(* IEC 61131-3 sources: krc-sample-programs/robot-cell-ethernetip-codesys/source/06_Programs, 5 files *)

(* ---- DASHBOARD.st ---- *)
PROGRAM DASHBOARD
VAR
	ipRobot      : NBS.IPv4Address := (ipAddress := ROBOT_IP);	// The robot's address
	fbClient     : NBS.TCP_Client;	// The connection to the robot's Dashboard Server
	fbWrite      : NBS.TCP_Write;	// Sends one line
	fbRead       : NBS.TCP_Read;	// Takes in whatever the robot has sent
	TON_POLL     : TON;	// Paces the questions
	TON_REPLY    : TON;	// The robot's answer is overdue
	TON_RETRY    : TON;	// Still not connected: try again
	bDropped     : BOOL;	// The connection was dropped this scan, so the retry timer starts over
	iDashStep    : INT;	// 0 not connected, 10 waiting for hello, 20 idle, 30 sending, 40 waiting for the answer
	bReconnect   : BOOL;	// Drop the connection for one scan, to connect again
	bAskRemote   : BOOL;	// The question in flight, or the next one, is remote control (the two take turns)
	sOut         : STRING(80);	// The line going out, with its line feed
	abIn         : ARRAY[0..127] OF BYTE;	// The bytes the read brings in
	sLine        : STRING(80);	// The line coming in, put together up to its line feed
	bLineDone    : BOOL;	// A whole line has come in this scan
	sChar        : STRING(1);	// One character, to add to the line
	i            : UDINT;	// Counts through the bytes read
END_VAR
// ---- body ----
// DASHBOARD: the driver for the second connection to the robot, its Dashboard Server. Not EtherNet/IP: one
// line of text over TCP to port 29999, and one line back. It asks the robot two questions, in turn, four times
// a second: what is the program doing ("programState": PLAYING, PAUSED, or STOPPED), and is the robot in
// remote control ("is in remote control": true or false). It leaves the answers in GVL_Link for INPUTS to read.
// (The Dashboard can also play, stop, and pause the program; here the register bits do that.)
// In simulation it doesn't run: SIM plays the robot's answers.
IF SIM_ENABLED THEN
    RETURN;
END_IF

// The connection: always on, except for the one scan it's dropped on purpose because the robot went quiet.
fbClient(xEnable := NOT bReconnect, itfIPAddress := ipRobot, uiPort := DASH_PORT);
bReconnect := FALSE;

// Take in what the robot sent, a byte at a time, until the line feed that ends its answer.
fbRead(xEnable := fbClient.xActive, itfConnection := fbClient.itfConnection, pData := ADR(abIn), udiSize := SIZEOF(abIn));
bLineDone := FALSE;
IF fbRead.xReady AND fbRead.udiCount > 0 THEN
    FOR i := 0 TO fbRead.udiCount - 1 DO
        IF abIn[i] = 10 THEN
            bLineDone := TRUE;
        ELSIF abIn[i] <> 13 AND LEN(sLine) < 80 THEN
            sChar[0] := abIn[i];
            sLine := CONCAT(sLine, sChar);
        END_IF
    END_FOR
END_IF

// Send the line, when there's one to send.
fbWrite(xExecute := iDashStep = 30, itfConnection := fbClient.itfConnection, pData := ADR(sOut), udiSize := INT_TO_UDINT(LEN(sOut)));

// The timers: one paces the questions, one gives up on an answer that doesn't come, and one on a connection that
// doesn't come (a refused or reset connection leaves the client in error until it is dropped and enabled again;
// on the bench, 2026-10-30, after the cable was out for minutes it never came back without this).
TON_POLL(IN := iDashStep = 20 AND NOT TON_POLL.Q, PT := DASH_POLL_TIME);
TON_REPLY(IN := iDashStep = 10 OR iDashStep = 40, PT := DASH_REPLY_TIME);
TON_RETRY(IN := iDashStep = 0 AND NOT fbClient.xActive AND NOT bDropped, PT := DASH_REPLY_TIME);
bDropped := FALSE;

CASE iDashStep OF
0:  // Not connected. When the connection comes up, the robot says hello first, and it can come in on the very
    // scan the connection does (it did on the bench, 2026-10-29): then it's already here, so don't wait for it.
    IF fbClient.xActive AND bLineDone THEN
        sLine := '';
        iDashStep := 20;
    ELSIF fbClient.xActive THEN
        iDashStep := 10;
    ELSE
        sLine := '';
    END_IF

10: // Waiting for hello: "Connected: Universal Robots Dashboard Server".
    IF bLineDone THEN
        sLine := '';
        iDashStep := 20;
    END_IF

20: // Idle. When it's time, the next question.
    IF TON_POLL.Q THEN
        bAskRemote := NOT bAskRemote;
        IF bAskRemote THEN
            sOut := 'is in remote control$N';
        ELSE
            sOut := 'programState$N';
        END_IF
        iDashStep := 30;
    END_IF

30: // Sending. When the line is out, wait for the answer.
    IF fbWrite.xDone THEN
        iDashStep := 40;
    END_IF
    IF fbWrite.xError THEN
        bReconnect := TRUE;
        iDashStep := 0;
    END_IF

40: // Waiting for the answer. Put it where it belongs.
    IF bLineDone THEN
        LINK_sDashReply := sLine;
        IF bAskRemote THEN
            LINK_bRemoteControl := sLine = 'true';
        ELSE
            LINK_sProgramState := sLine;
        END_IF
        sLine := '';
        iDashStep := 20;
    END_IF
END_CASE

// The robot went quiet, or never answered the call: drop the connection and connect again.
IF TON_REPLY.Q OR TON_RETRY.Q THEN
    bReconnect := TRUE;
    bDropped := TRUE;
    iDashStep := 0;
END_IF

// Without the connection, nothing the robot said last still counts.
IF NOT fbClient.xActive THEN
    iDashStep := 0;
    LINK_sProgramState := '';
    LINK_bRemoteControl := FALSE;
END_IF
LINK_bDashConnected := fbClient.xActive AND iDashStep >= 20;

(* ---- DEVICES.st ---- *)
PROGRAM DEVICES
VAR
	iDeviceStep : E_Step;	// The step the devices follow: the step itself, or while paused, the step Pause came from
END_VAR
// ---- body ----
// DEVICES: every output is set here, once, from the step. Nothing here reads a button or another output.
// Each bit is written like a coil: TRUE while its condition is true, FALSE as soon as it isn't.

// While paused, the clamp, the command, and fixture clear stay as they were in the step Pause came from,
// so the robot carries on where it left off and a clamped part stays clamped.
IF iStep = S9_PAUSED OR iStep = S9_RESUMING THEN
    iDeviceStep := iPausedStep;
ELSE
    iDeviceStep := iStep;
END_IF

// Command to the robot: load in the two load steps, unload in the two unload steps, 0 everywhere else.
// Clearing it is the PLC's half of ending a handshake.
IF iDeviceStep = S4_LOAD_REQUEST OR iDeviceStep = S4_LOADING THEN
    diCommand := CMD_LOAD;
ELSIF iDeviceStep = S7_UNLOAD_REQUEST OR iDeviceStep = S7_UNLOADING THEN
    diCommand := CMD_UNLOAD;
ELSE
    diCommand := CMD_NONE;
END_IF

// Fixture clear: the robot may reach into the fixture, only while it's loading or unloading and the
// clamp reads open. The robot program waits for it before it goes in.
bFixtureClear := (iDeviceStep = S4_LOAD_REQUEST OR iDeviceStep = S4_LOADING OR iDeviceStep = S7_UNLOAD_REQUEST
    OR iDeviceStep = S7_UNLOADING) AND bClampOpen;

// The robot program's Start, Stop, and Pause: three register bits the robot has set up as I/O actions. Each
// acts as its bit turns on: Start while starting or resuming, Stop in Stopped, Pause in Paused.
bRobotStart := iStep = S3_STARTING OR iStep = S9_RESUMING;
bRobotStop := iStep = S8_STOPPED;
bRobotPause := iStep = S9_PAUSED;

// PLC heartbeat: counted up every 250 ms, in every step, so the robot can tell the PLC is still running.
// The timer restarts itself each time it fires.
TON_PLC_BEAT(IN := NOT TON_PLC_BEAT.Q, PT := HEARTBEAT_TIME);
IF TON_PLC_BEAT.Q THEN
    diPlcHeartbeat := diPlcHeartbeat + 1;
END_IF

// Clamp valve: on in Clamping and Holding.
bClampClose := iDeviceStep = S5_CLAMPING OR iDeviceStep = S5_HOLDING;

// Pressure setpoint to the regulator: the HMI setpoint while the valve is on, 0 the rest of the time.
IF iDeviceStep = S5_CLAMPING OR iDeviceStep = S5_HOLDING THEN
    rPressureSet := HMI_rPressureSet;
ELSE
    rPressureSet := 0.0;
END_IF

// Stack light green: ready, starting, cycling, or paused (the cycle is on hold, nothing is wrong).
bStackGreen := (iStep >= S3_READY AND iStep <= S7_UNLOAD_CLEAR) OR iStep = S9_PAUSED OR iStep = S9_RESUMING;

// Stack light red: not ready to cycle. Written from the steps, never as "not green".
bStackRed := iStep = S0_IDLE OR iStep = S1_NOT_READY OR iStep = S2_RESET OR iStep = S8_FAULT OR iStep = S8_STOPPED;

// Stack light orange: faulted.
bStackOrange := iStep = S8_FAULT;

// Start lamp: lit when Start does something: in Ready, and in Paused once the robot program has paused.
// Everywhere else Start does nothing.
bStartLamp := iStep = S3_READY OR (iStep = S9_PAUSED AND bProgramPaused);

// Stop lamp: lit when Stop does something, everywhere but Stopped.
bStopLamp := iStep <> S8_STOPPED;

// Pause lamp: lit when Pause does something, in a cycle.
bPauseLamp := iStep >= S4_LOAD_REQUEST AND iStep <= S7_UNLOAD_CLEAR;

// Reset lamp: lit when the cell is faulted or stopped and needs a reset.
bResetLamp := iStep = S8_FAULT OR iStep = S8_STOPPED;

(* ---- INPUTS.st ---- *)
// SAMPLE PROGRAM: a clamp station loaded and unloaded by a robot. KRC (Kurtin Robotics), written as a teaching
// example. The PLC (WAGO CC100) runs the cell and talks to a Universal Robots arm over EtherNet/IP: it tells the
// robot to load a part, clamps it to a pressure setpoint from the HMI, holds, opens, and tells the robot to
// unload it. Every command is a handshake (command, acknowledge, done, clear), every step of it has a timeout,
// and the PLC watches the robot's heartbeat. The panel's Start, Stop, and Pause work the robot program through
// three register bits, and a second connection, the robot's Dashboard, tells the PLC whether the program is
// playing, paused, or stopped. Each fault says which side failed.
// NOT A SAFETY FUNCTION. Nothing on this link stops the robot. Stopping motion is the robot's safety system
// (its protective and emergency stops); the PLC only watches it.
// How it is laid out: MainTask calls SIM (simulation only), then INPUTS, STATE_MACHINE, DEVICES, OUTPUTS, and
// DASHBOARD, every scan. INPUTS reads every input, the robot's words included, into a program tag. STATE_MACHINE
// decides the step. DEVICES sets every output from the step. OUTPUTS writes every output to the hardware, the
// robot, and the HMI. DASHBOARD is the driver for the Dashboard connection: it asks the robot what its program
// is doing.
PROGRAM INPUTS
// ---- body ----
// INPUTS: every input is read here and nowhere else.
// Start: the panel button or the HMI button. The state machine acts on the press, the scan it goes on, so
// a button held down (or stuck) can't start one cycle after another.
bStartPB := DI_bStartPB OR HMI_bStartPB;
bStartPressed := bStartPB AND NOT bStartLast;
bStartLast := bStartPB;

// Stop is wired normally closed: the input is on while nobody presses it, so a broken wire reads the
// same as pressing Stop. This is the only place it gets turned around. Or the Stop button on the HMI.
bStopPB := NOT DI_bStopPB_NC OR HMI_bStopPB;

// Reset: the panel button or the HMI button.
bResetPB := DI_bResetPB OR HMI_bResetPB;

// Pause: the HMI button.
bPausePB := HMI_bPausePB;

// The clamp open sensor and the part-present sensor in the fixture.
bClampOpen := DI_bClampOpen;
bPartPresent := DI_bPartPresent;

// Pressure: the CC100 reads 0 to 10 V as 0 to 32760. Scaled once, here, to psi.
rPressure := WORD_TO_REAL(AI_wPressure) * PRESSURE_RANGE / AI_FULL_SCALE;

// The link's own health. On a real controller it's the scanner's word on the robot's connection, from the
// robot's device, UR_Robot. In simulation the scanner doesn't run, so SIM plays it instead.
IF NOT SIM_ENABLED THEN
    LINK_bCommError := UR_Robot.State <> IoDrvEtherNetIP.ADAPTERSTATE.RUNNING;
END_IF
bLinkError := LINK_bCommError;

// The robot's words, read once, each into a tag with a name.
diRobotHeartbeat := LINK_adiFromRobot[FROM_HEARTBEAT];
bRobotReady := LINK_adiFromRobot[FROM_READY] = 1;
diRobotAck := LINK_adiFromRobot[FROM_ACK];
diRobotDone := LINK_adiFromRobot[FROM_DONE];
diRobotFault := LINK_adiFromRobot[FROM_FAULT];
diRobotStep := LINK_adiFromRobot[FROM_ROBOT_STEP];
bHandshakeClear := diRobotAck = CMD_NONE AND diRobotDone = CMD_NONE;

// The robot controller's own state, from the same EtherNet/IP assembly: its mode, whether its program is
// running, and its stops (a safeguard stop is a protective stop from a guard; the three emergency stops are
// the system's, the robot's, and the cell's).
bRobotRunning := LINK_siRobotMode = ROBOT_RUNNING;
bProgramRunning := LINK_dwRobotBits.1;
bRobotProtStop := LINK_dwSafetyBits.2 OR LINK_dwSafetyBits.4;
bRobotEStop := LINK_dwSafetyBits.5 OR LINK_dwSafetyBits.6 OR LINK_dwSafetyBits.7;

// The Dashboard's answers: the connection, whether the robot program is playing, paused, or stopped (all
// EtherNet/IP can say is running or not), and whether the robot is in remote control.
bDashConnected := LINK_bDashConnected;
bProgramPlaying := FIND(LINK_sProgramState, 'PLAYING') = 1;
bProgramPaused := FIND(LINK_sProgramState, 'PAUSED') = 1;
bProgramStopped := FIND(LINK_sProgramState, 'STOPPED') = 1;
bRemoteControl := LINK_bRemoteControl;

// The robot's heartbeat: its program counts it up. If the count hasn't changed for a second, the robot
// program has stopped. The timer only runs while the count stands still, so every change restarts it.
TON_BEAT_LOST(IN := diRobotHeartbeat = diRobotBeatLast, PT := HEARTBEAT_LOST);
bRobotAlive := NOT TON_BEAT_LOST.Q;
diRobotBeatLast := diRobotHeartbeat;

// The timeouts from the HMI, in seconds, as each timer's preset.
TON_ACK.PT := T#1S * HMI_iAckTimeout;
TON_CLEAR.PT := T#1S * HMI_iAckTimeout;
TON_MOVE.PT := T#1S * HMI_iMoveTimeout;
TON_CLAMP.PT := T#1S * HMI_iClampTimeout;
TON_HOLD.PT := T#1S * HMI_iHoldTime;
TON_OPEN.PT := T#1S * HMI_iOpenTimeout;

(* ---- OUTPUTS.st ---- *)
PROGRAM OUTPUTS
// ---- body ----
// OUTPUTS: every output is written here and nowhere else. First the hardware, in terminal order.
DO_bClampClose := bClampClose;
DO_bStackGreen := bStackGreen;
DO_bStackRed := bStackRed;
DO_bStackOrange := bStackOrange;

// Pressure setpoint to the regulator: the input's scaling, run backwards. 0 to 32767 for 0 to 10 V.
AO_wPressureSet := REAL_TO_WORD(rPressureSet * AO_FULL_SCALE / PRESSURE_RANGE);

// Then the robot: the four words to its input registers 0 to 3, sent every EtherNet/IP cycle.
LINK_adiToRobot[TO_HEARTBEAT] := diPlcHeartbeat;
LINK_adiToRobot[TO_COMMAND] := diCommand;
LINK_adiToRobot[TO_FIXTURE_CLEAR] := BOOL_TO_DINT(bFixtureClear);
LINK_adiToRobot[TO_PLC_STEP] := INT_TO_DINT(iStep);

// And the robot program's Start, Stop, and Pause bits, input bit registers 0 to 2.
LINK_dwToRobotBits.BIT_START := bRobotStart;
LINK_dwToRobotBits.BIT_STOP := bRobotStop;
LINK_dwToRobotBits.BIT_PAUSE := bRobotPause;

// Then the HMI. The screen only reads these.
HMI_bStartLamp := bStartLamp;
HMI_bStopLamp := bStopLamp;
HMI_bResetLamp := bResetLamp;
HMI_bPauseLamp := bPauseLamp;
HMI_bStackGreen := bStackGreen;
HMI_bStackRed := bStackRed;
HMI_bStackOrange := bStackOrange;
HMI_rPressure := rPressure;
HMI_sState := sStateDescription;
HMI_bLinkUp := NOT bLinkError AND bRobotAlive;
HMI_bDashUp := bDashConnected;
HMI_bRemote := bRemoteControl;
HMI_bProgramRunning := bProgramRunning;
HMI_bRobotReady := bRobotReady;
HMI_bRobotRunning := bRobotRunning;
HMI_bRobotStopped := bRobotProtStop OR bRobotEStop;
HMI_bPartPresent := bPartPresent;
HMI_iToRobot[0] := LINK_adiToRobot[0];
HMI_iToRobot[1] := LINK_adiToRobot[1];
HMI_iToRobot[2] := LINK_adiToRobot[2];
HMI_iToRobot[3] := LINK_adiToRobot[3];
HMI_iToRobot[4] := DWORD_TO_DINT(LINK_dwToRobotBits AND 16#7);
HMI_iFromRobot[0] := LINK_adiFromRobot[0];
HMI_iFromRobot[1] := LINK_adiFromRobot[1];
HMI_iFromRobot[2] := LINK_adiFromRobot[2];
HMI_iFromRobot[3] := LINK_adiFromRobot[3];
HMI_iFromRobot[4] := LINK_adiFromRobot[4];
HMI_iFromRobot[5] := LINK_adiFromRobot[5];

// What the robot program is doing, in words, from the step it writes as it goes. The step only means
// something while the program plays: stopped or paused, the register still holds the last step written.
IF NOT bDashConnected THEN
    HMI_sRobot := 'Robot: no Dashboard connection';
ELSIF bProgramPaused THEN
    HMI_sRobot := 'Robot: program paused';
ELSIF NOT bProgramRunning AND diRobotStep = ROBOT_NOT_HOME THEN
    HMI_sRobot := 'Robot: started away from home and stopped, jog it home';
ELSIF NOT bProgramRunning THEN
    HMI_sRobot := 'Robot: program stopped';
ELSE
    CASE diRobotStep OF
    10:  HMI_sRobot := 'Robot: starting, checking it is at home';
    100: HMI_sRobot := 'Robot: at home, waiting for a command';
    200: HMI_sRobot := 'Robot: load, picking a part';
    210: HMI_sRobot := 'Robot: load, waiting for fixture clear';
    220: HMI_sRobot := 'Robot: load, placing the part';
    300: HMI_sRobot := 'Robot: unload, waiting for fixture clear';
    310: HMI_sRobot := 'Robot: unload, taking the part out';
    320: HMI_sRobot := 'Robot: unload, dropping the part';
    400: HMI_sRobot := 'Robot: done, waiting for the PLC to clear the command';
    800: HMI_sRobot := 'Robot: gripper missed, going home';
    ELSE
        HMI_sRobot := CONCAT('Robot: step ', DINT_TO_STRING(diRobotStep));
    END_CASE
END_IF

(* ---- STATE_MACHINE.st ---- *)
PROGRAM STATE_MACHINE
VAR
	bAllClear  : BOOL;	// Everything the cell needs before it can be Ready
	bCycling   : BOOL;	// The cell is in a cycle, from Load request to Unload clear
	bRobotBusy : BOOL;	// The robot program has work from the PLC: starting, cycling, paused, or resuming
END_VAR
// ---- body ----
// STATE_MACHINE: decides which step the cell is in. One CASE on the step, one branch per step.
// Inside a branch, each exit is one IF: the reason it leaves, then the next step into iNextStep and what
// the cell will be doing, for the HMI. The step only changes on the last line, so every line in one
// scan sees the same step.

// The step timers. Each runs only while its steps are active, so it starts from zero every time.
TON_START(IN := iStep = S3_STARTING OR iStep = S9_RESUMING, PT := ROBOT_START_TIME);
TON_PAUSE(IN := iStep = S9_PAUSED AND NOT bProgramPaused, PT := ROBOT_PAUSE_TIME);
TON_ACK(IN := iStep = S4_LOAD_REQUEST OR iStep = S7_UNLOAD_REQUEST);
TON_MOVE(IN := iStep = S4_LOADING OR iStep = S7_UNLOADING);
TON_CLEAR(IN := iStep = S4_LOAD_CLEAR OR iStep = S7_UNLOAD_CLEAR);
TON_CLAMP(IN := iStep = S5_CLAMPING);
TON_HOLD(IN := iStep = S5_HOLDING);
TON_OPEN(IN := iStep = S6_OPENING);

// Everything the cell needs before it's Ready: the link up, the Dashboard up and the robot in remote control
// (so it takes Start, Stop, and Pause), the arm Running with no stop on it, the robot program not paused, and
// if it's already running, its heartbeat ticking, ready, and the last handshake cleared; the clamp open, the
// fixture empty, and Stop not pressed. A stopped robot program is fine: Start starts it.
bAllClear := NOT bLinkError AND bDashConnected AND bRemoteControl AND bRobotRunning AND NOT bRobotProtStop
    AND NOT bRobotEStop AND NOT bProgramPaused
    AND (NOT bProgramRunning OR (bRobotAlive AND bRobotReady AND bHandshakeClear))
    AND bClampOpen AND NOT bPartPresent AND NOT bStopPB;
bCycling := iStep >= S4_LOAD_REQUEST AND iStep <= S7_UNLOAD_CLEAR;
bRobotBusy := bCycling OR iStep = S3_STARTING OR iStep = S9_PAUSED OR iStep = S9_RESUMING;

CASE iStep OF

S0_IDLE:
    // Idle: powered up and at rest. Go to Not Ready.
    iNextStep := S1_NOT_READY;
    sStateDescription := 'Not Ready - waiting for the robot and an empty fixture';

S1_NOT_READY:
    // Not Ready: all clear. Ready.
    IF bAllClear THEN
        iNextStep := S3_READY;
        sStateDescription := 'Ready - press Start';
    END_IF
    // Not Ready: Reset pressed. Go through Reset.
    IF bResetPB THEN
        iNextStep := S2_RESET;
        sStateDescription := 'Reset - release Reset';
    END_IF

S2_RESET:
    // Reset: Reset released. Back to Not Ready, which checks everything again before Ready.
    IF NOT bResetPB THEN
        iNextStep := S1_NOT_READY;
        sStateDescription := 'Not Ready - waiting for the robot and an empty fixture';
    END_IF

S3_READY:
    // Ready: Start pressed (just now, not held) and the robot program isn't running. Start it.
    IF bStartPressed AND NOT bProgramRunning THEN
        iNextStep := S3_STARTING;
        sStateDescription := 'Starting - starting the robot program';
    END_IF
    // Ready: Start pressed and the robot program is already running. Ask it to load a part.
    IF bStartPressed AND bProgramRunning THEN
        iNextStep := S4_LOAD_REQUEST;
        sStateDescription := 'Load - asking the robot to load a part';
    END_IF
    // Ready: anything in all clear is gone (the robot dropped out). Back to Not Ready. Written last, so it wins.
    IF NOT bAllClear THEN
        iNextStep := S1_NOT_READY;
        sStateDescription := 'Not Ready - waiting for the robot and an empty fixture';
    END_IF

S3_STARTING:
    // Starting: the robot program runs, its heartbeat ticks, and it's at home, ready. Ask it to load a part.
    IF bProgramRunning AND bRobotAlive AND bRobotReady AND bHandshakeClear THEN
        iNextStep := S4_LOAD_REQUEST;
        sStateDescription := 'Load - asking the robot to load a part';
    END_IF
    // Starting: not running and ready in time. Fault, on the robot's side.
    IF TON_START.Q THEN
        iNextStep := S8_FAULT;
        sStateDescription := 'Fault - robot program did not start in time';
    END_IF
    // Starting: the robot program found itself away from home and stopped rather than move. Given time to
    // start and write its step first, so an old step from last time doesn't count. Written last, so it wins.
    IF TON_START.ET >= ROBOT_HOME_CHECK AND diRobotStep = ROBOT_NOT_HOME AND NOT bProgramRunning THEN
        iNextStep := S8_FAULT;
        sStateDescription := 'Fault - robot is away from home, jog it home';
    END_IF

S4_LOAD_REQUEST:
    // Load request: the robot echoes the load command. It's on its way.
    IF diRobotAck = CMD_LOAD THEN
        iNextStep := S4_LOADING;
        sStateDescription := 'Load - the robot is loading a part';
    END_IF
    // Load request: no answer in time. Fault, on the robot's side.
    IF TON_ACK.Q AND diRobotAck <> CMD_LOAD THEN
        iNextStep := S8_FAULT;
        sStateDescription := 'Fault - robot did not acknowledge the load';
    END_IF

S4_LOADING:
    // Loading: the robot says done and the fixture sees the part. Clear the handshake.
    IF diRobotDone = CMD_LOAD AND bPartPresent THEN
        iNextStep := S4_LOAD_CLEAR;
        sStateDescription := 'Load - part in, clearing the handshake';
    END_IF
    // Loading: the robot says done but the fixture doesn't see a part. Fault, checked on the PLC's side.
    IF diRobotDone = CMD_LOAD AND NOT bPartPresent THEN
        iNextStep := S8_FAULT;
        sStateDescription := 'Fault - robot finished the load but no part in the fixture';
    END_IF
    // Loading: no done in time. Fault, on the robot's side.
    IF TON_MOVE.Q AND diRobotDone <> CMD_LOAD THEN
        iNextStep := S8_FAULT;
        sStateDescription := 'Fault - robot did not finish the load in time';
    END_IF
    // Loading: the robot reports its own fault. Written last, so it wins.
    IF diRobotFault <> 0 THEN
        iNextStep := S8_FAULT;
        sStateDescription := 'Fault - robot reports its gripper missed the part';
    END_IF

S4_LOAD_CLEAR:
    // Load clear: the robot cleared its acknowledge and done. Clamp the part.
    IF bHandshakeClear THEN
        iNextStep := S5_CLAMPING;
        sStateDescription := 'Clamping - building pressure';
    END_IF
    // Load clear: the robot didn't clear in time. Fault, on the robot's side.
    IF TON_CLEAR.Q AND NOT bHandshakeClear THEN
        iNextStep := S8_FAULT;
        sStateDescription := 'Fault - robot did not clear the handshake';
    END_IF

S5_CLAMPING:
    // Clamping: the pressure is within the band of the setpoint. Hold it.
    IF rPressure >= HMI_rPressureSet - PRESSURE_BAND THEN
        iNextStep := S5_HOLDING;
        sStateDescription := 'Clamping - holding at pressure';
    END_IF
    // Clamping: the timeout ran out and the pressure is still short. Fault, on the clamp.
    IF TON_CLAMP.Q AND rPressure < HMI_rPressureSet - PRESSURE_BAND THEN
        iNextStep := S8_FAULT;
        sStateDescription := 'Fault - pressure not reached in time';
    END_IF

S5_HOLDING:
    // Holding: the hold time is up. Open the clamp.
    IF TON_HOLD.Q THEN
        iNextStep := S6_OPENING;
        sStateDescription := 'Opening - hold done';
    END_IF

S6_OPENING:
    // Opening: the clamp reads open. Ask the robot to unload the part.
    IF bClampOpen THEN
        iNextStep := S7_UNLOAD_REQUEST;
        sStateDescription := 'Unload - asking the robot to unload the part';
    END_IF
    // Opening: the timeout ran out and the clamp still doesn't read open. Fault, on the clamp.
    IF TON_OPEN.Q AND NOT bClampOpen THEN
        iNextStep := S8_FAULT;
        sStateDescription := 'Fault - clamp did not open in time';
    END_IF

S7_UNLOAD_REQUEST:
    // Unload request: the robot echoes the unload command. It's on its way.
    IF diRobotAck = CMD_UNLOAD THEN
        iNextStep := S7_UNLOADING;
        sStateDescription := 'Unload - the robot is unloading the part';
    END_IF
    // Unload request: no answer in time. Fault, on the robot's side.
    IF TON_ACK.Q AND diRobotAck <> CMD_UNLOAD THEN
        iNextStep := S8_FAULT;
        sStateDescription := 'Fault - robot did not acknowledge the unload';
    END_IF

S7_UNLOADING:
    // Unloading: the robot says done and the fixture is empty. Clear the handshake.
    IF diRobotDone = CMD_UNLOAD AND NOT bPartPresent THEN
        iNextStep := S7_UNLOAD_CLEAR;
        sStateDescription := 'Unload - part out, clearing the handshake';
    END_IF
    // Unloading: the robot says done but the part is still in the fixture. Fault, checked on the PLC's side.
    IF diRobotDone = CMD_UNLOAD AND bPartPresent THEN
        iNextStep := S8_FAULT;
        sStateDescription := 'Fault - robot finished the unload but the part is still in the fixture';
    END_IF
    // Unloading: no done in time. Fault, on the robot's side.
    IF TON_MOVE.Q AND diRobotDone <> CMD_UNLOAD THEN
        iNextStep := S8_FAULT;
        sStateDescription := 'Fault - robot did not finish the unload in time';
    END_IF
    // Unloading: the robot reports its own fault. Written last, so it wins.
    IF diRobotFault <> 0 THEN
        iNextStep := S8_FAULT;
        sStateDescription := 'Fault - robot reports its gripper missed the part';
    END_IF

S7_UNLOAD_CLEAR:
    // Unload clear, single cycle: the robot cleared its answer. The part is done: Ready for the next Start.
    IF bHandshakeClear AND NOT HMI_bContinuous THEN
        iNextStep := S3_READY;
        sStateDescription := 'Ready - press Start';
    END_IF
    // Unload clear, continuous: the part is done, straight into the next one, until Stop or Pause (or the
    // switch back to single cycle, which finishes this part and stops at Ready).
    IF bHandshakeClear AND HMI_bContinuous THEN
        iNextStep := S4_LOAD_REQUEST;
        sStateDescription := 'Load - asking the robot to load a part';
    END_IF
    // Unload clear: the robot didn't clear in time. Fault, on the robot's side.
    IF TON_CLEAR.Q AND NOT bHandshakeClear THEN
        iNextStep := S8_FAULT;
        sStateDescription := 'Fault - robot did not clear the handshake';
    END_IF

S8_FAULT:
    // Fault: Reset pressed. Go through Reset, then Not Ready.
    IF bResetPB THEN
        iNextStep := S2_RESET;
        sStateDescription := 'Reset - release Reset';
    END_IF

S8_STOPPED:
    // Stopped: Stop released and Reset pressed. Go through Reset, then Not Ready.
    IF bResetPB AND NOT bStopPB THEN
        iNextStep := S2_RESET;
        sStateDescription := 'Reset - release Reset';
    END_IF

S9_PAUSED:
    // Paused: the Dashboard says the robot program is paused, and Start is pressed. Carry on.
    IF bStartPressed AND bProgramPaused THEN
        iNextStep := S9_RESUMING;
        sStateDescription := 'Paused - resuming the robot program';
    END_IF
    // Paused: the robot program never paused. Fault, on the robot's side.
    IF TON_PAUSE.Q AND NOT bProgramStopped THEN
        iNextStep := S8_FAULT;
        sStateDescription := 'Fault - robot program did not pause';
    END_IF
    // Paused: the Dashboard says the robot program is stopped, not paused (stopped on the pendant, or it hit
    // an error). Start would run it from the top, not carry on, so the cycle can't go on. Fault. Written
    // last, so it wins.
    IF bProgramStopped THEN
        iNextStep := S8_FAULT;
        sStateDescription := 'Fault - robot program stopped while paused, it cannot carry on';
    END_IF

S9_RESUMING:
    // Resuming: the robot program runs and its heartbeat ticks. Back to the step Pause came from.
    IF bProgramRunning AND bRobotAlive THEN
        iNextStep := iPausedStep;
        sStateDescription := sPausedDescription;
    END_IF
    // Resuming: not running in time. Fault, on the robot's side.
    IF TON_START.Q THEN
        iNextStep := S8_FAULT;
        sStateDescription := 'Fault - robot program did not resume in time';
    END_IF
END_CASE

// Pause, in a cycle: remember where the cycle was going and what it was doing, and pause. Only while that
// is still a cycle step (an exit above may already be a fault, or the end of the cycle).
IF bCycling AND bPausePB AND iNextStep >= S4_LOAD_REQUEST AND iNextStep <= S7_UNLOAD_CLEAR THEN
    iPausedStep := iNextStep;
    sPausedDescription := sStateDescription;
    iNextStep := S9_PAUSED;
    sStateDescription := 'Paused - press Start to carry on';
END_IF

// While the robot has work, losing the robot wins over every exit above. Each has its own words, so the
// screen says which side failed. Written in this order, so the last true one wins: the arm stops Running,
// the robot's heartbeat stops (its program stopped; only checked in a cycle, since a paused or starting
// program doesn't count), the robot leaves remote control, the Dashboard drops, its protective stop, its
// emergency stop, and last the network, because with the link down every word from the robot is stale.
IF bRobotBusy AND NOT bRobotRunning THEN
    iNextStep := S8_FAULT;
    sStateDescription := 'Fault - robot arm not running';
END_IF
IF bCycling AND NOT bRobotAlive THEN
    iNextStep := S8_FAULT;
    sStateDescription := 'Fault - no robot heartbeat, robot program stopped';
END_IF
IF bRobotBusy AND bDashConnected AND NOT bRemoteControl THEN
    iNextStep := S8_FAULT;
    sStateDescription := 'Fault - robot left remote control';
END_IF
IF bRobotBusy AND NOT bDashConnected THEN
    iNextStep := S8_FAULT;
    sStateDescription := 'Fault - Dashboard connection lost';
END_IF
IF bRobotBusy AND bRobotProtStop THEN
    iNextStep := S8_FAULT;
    sStateDescription := 'Fault - robot in a protective stop';
END_IF
IF bRobotBusy AND bRobotEStop THEN
    iNextStep := S8_FAULT;
    sStateDescription := 'Fault - robot emergency stop';
END_IF
IF bRobotBusy AND bLinkError THEN
    iNextStep := S8_FAULT;
    sStateDescription := 'Fault - link lost, PLC cannot reach the robot';
END_IF

// Stop, from any step: the robot program stops right away and the cell waits in Stopped for Reset. It's
// the operator's word, so it wins over everything. (Stop is not a safety function: stopping the robot for
// a person is its own safety system.)
IF bStopPB AND iStep <> S8_STOPPED THEN
    iNextStep := S8_STOPPED;
    sStateDescription := 'Stopped - robot program stopped, press Reset';
END_IF

// Take the next step. This is the only place the step changes.
iStep := iNextStep;
